// TIA Portal V21 export
VAR_GLOBAL   // PLC tag table "Signalläuchte"
   LED_rot AT %Q1.4 : Bool;
   LED_gelb AT %Q1.6 : Bool;
   LED_grün AT %Q1.5 : Bool;
END_VAR
